(* IEC 61131-3 sources: plc-st-coding-agent/progress/evidence/f14_v5_preflight_20261112, 2 files *)

(* ---- negative.st ---- *)
TYPE ST_V5_Probe : STRUCT value : INT; END_STRUCT END_TYPE;
FUNCTION_BLOCK FB_V5Probe
VAR_INPUT go:BOOL; mode:INT; END_VAR
VAR_OUTPUT rec:ST_V5_Probe; END_VAR
VAR state:(STATE_IDLE,STATE_ACTIVE); END_VAR
IF go THEN state:=STATE_ACTIVE; END_IF;
CASE mode OF
1: IF go THEN
CASE state OF
STATE_IDLE: rec.value:=3;
STATE_ACTIVE: undeclared_v5_bad:=7;
END_CASE;
END_IF;
2: rec.value:=9;
END_CASE;
END_FUNCTION_BLOCK

(* ---- positive.st ---- *)
TYPE ST_V5_Probe : STRUCT value : INT; END_STRUCT END_TYPE;
FUNCTION_BLOCK FB_V5Probe
VAR_INPUT go:BOOL; mode:INT; END_VAR
VAR_OUTPUT rec:ST_V5_Probe; END_VAR
VAR state:(STATE_IDLE,STATE_ACTIVE); END_VAR
IF go THEN state:=STATE_ACTIVE; END_IF;
CASE mode OF
1: IF go THEN
CASE state OF
STATE_IDLE: rec.value:=3;
STATE_ACTIVE: rec.value:=7;
END_CASE;
END_IF;
2: rec.value:=9;
END_CASE;
END_FUNCTION_BLOCK
